// TIA Portal V19 export
FUNCTION_BLOCK "HEATING_PROCEES"   // FB14, LAD
TITLE = Heating
{ S7_Optimized_Access := 'TRUE' }
// stored: MemoryReserve 100, SetENOAutomatically false
   VAR_INPUT
      CHS_CFB : Bool;
      UCHS_CFB : Bool;
      CSV_CFB : Bool;
      HEAT_RUNNING : Bool;
      SELECT_CHWS : Bool;
      SELECT_CTS : Bool;
      SELECT_HWS : Bool;
      RUNNING : Bool;
      ESTOP : Bool;
      RESET : Bool;
      UCHWS : Bool;
      CHWS : Bool;
      CTS : Bool;
      HWS : Bool;
      HWS_OFB : Bool;
      CTS_OFB : Bool;
      CHWS_OFB : Bool;
      PUMP_RUN : Bool;
      SP : Real;
      PV : Real;
   END_VAR
   VAR_OUTPUT
      UCHWS_CMD : Bool;
      UCHWR_CMD : Bool;
      CHWS_CMD : Bool;
      CHWR_CMD : Bool;
      CTS_CMD : Bool;
      CTR_CMD : Bool;
      HWS_CMD : Bool;
      HWR_CMD : Bool;
      PUMP_CMD : Bool;
      CV_CMD : Bool;
   END_VAR
   VAR
      IEC_Timer_0_Instance : TP_TIME;
      IEC_Timer_1_Instance_1 { S7_SetPoint := 'True'} : TP_TIME;
      IEC_Timer_0_Instance_1 { S7_SetPoint := 'True'} : TP_TIME;
      IEC_Timer_0_Instance_2 { S7_SetPoint := 'True'} : TP_TIME;
      IEC_Timer_0_Instance_3 { S7_SetPoint := 'True'} : TP_TIME;
      IEC_Timer_0_Instance_4 { S7_SetPoint := 'True'} : TP_TIME;
      IEC_Timer_0_Instance_5 { S7_SetPoint := 'True'} : TP_TIME;
      IEC_Timer_0_Instance_6 { S7_SetPoint := 'True'} : TP_TIME;
      IEC_Timer_0_Instance_7 { S7_SetPoint := 'True'} : TP_TIME;
      IEC_Timer_0_Instance_8 { S7_SetPoint := 'True'} : TP_TIME;
      IEC_Timer_0_Instance_9 { S7_SetPoint := 'True'} : TP_TIME;
      "STEP" { S7_SetPoint := 'True'} : Int;
      P_TRIG : Bool;
      P_TRIG_1 : Bool;
      P_TRIG_2 : Bool;
      P_TRIG_3 : Bool;
      P_TRIG_4 : Bool;
      P_TRIG_5 : Bool;
      P_TRIG_6 : Bool;
      P_TRIG_7 : Bool;
      P_TRIG_8 : Bool;
      P_TRIG_9 : Bool;
      P_TRIG_10 : Bool;
      P_TRIG_11 : Bool;
      P_TRIG_12 : Bool;
      P_TRIG_13 : Bool;
      P_TRIG_14 : Bool;
      P_TRIG_15 : Bool;
      P_TRIG_16 : Bool;
      IEC_Timer_0_Instance_10 { S7_SetPoint := 'True'} : TP_TIME;
      IEC_Timer_0_Instance_11 { S7_SetPoint := 'True'} : TON_TIME;
      IEC_Timer_0_Instance_12 { S7_SetPoint := 'True'} : TON_TIME;
   END_VAR
   VAR_TEMP   // added for the SCL form of the ladder/FBD networks
      _w1 : Bool;
      _w2 : Bool;
      _w3 : Bool;
      _w4 : Bool;
      _w5 : Bool;
      _w6 : Bool;
      _w7 : Bool;
      _w8 : Bool;
   END_VAR
BEGIN

REGION Network 1: ULTRACHILLED TO CHILLED MODE
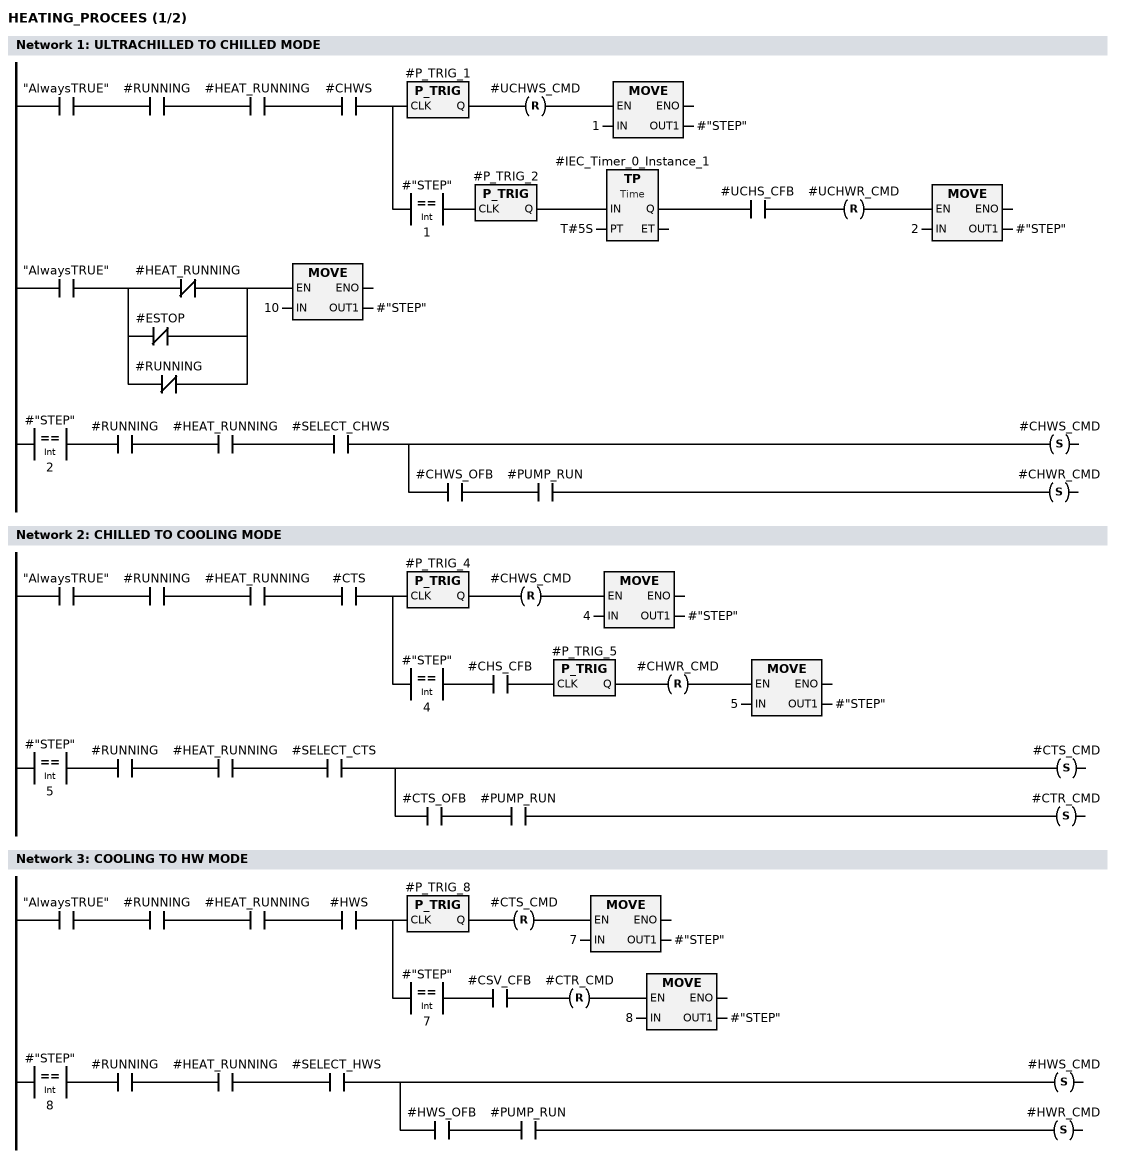
   RUNG wire#powerrail
      Contact( "AlwaysTRUE" )
      Contact( #RUNNING )
      Contact( #HEAT_RUNNING )
      Contact( #CHWS )
      wire#w1
      P_Trig( #P_TRIG_1 )
      R_Coil( #UCHWS_CMD )
      Move(in := 1, out1 => #"STEP")
   END_RUNG
   RUNG wire#w1
      { S7_Templates := "SrcType := Int" } EQ_Contact(in1 := #"STEP", in2 := 1)
      P_Trig( #P_TRIG_2 )
      { S7_Templates := "time_type := Time" } #IEC_Timer_0_Instance_1.TP(pt := T#5S, et =>)
      Contact( #UCHS_CFB )
      R_Coil( #UCHWR_CMD )
      Move(in := 2, out1 => #"STEP")
   END_RUNG
   RUNG wire#powerrail
      Contact( "AlwaysTRUE" )
      wire#w2
      I_Contact( #HEAT_RUNNING )
      wire#w3
      Move(in := 10, out1 => #"STEP")
   END_RUNG
   RUNG wire#w2
      I_Contact( #ESTOP )
   END_RUNG wire#w3
   RUNG wire#w2
      I_Contact( #RUNNING )
   END_RUNG wire#w3
   RUNG wire#powerrail
      { S7_Templates := "SrcType := Int" } EQ_Contact(in1 := #"STEP", in2 := 2)
      Contact( #RUNNING )
      Contact( #HEAT_RUNNING )
      Contact( #SELECT_CHWS )
      wire#w4
      S_Coil( #CHWS_CMD )
   END_RUNG
   RUNG wire#w4
      Contact( #CHWS_OFB )
      Contact( #PUMP_RUN )
      S_Coil( #CHWR_CMD )
   END_RUNG
   // the same network as SCL:
   #_w1 := "AlwaysTRUE" AND #RUNNING AND #HEAT_RUNNING AND #CHWS;
   #_w2 := #_w1 AND NOT #P_TRIG_1;   // rising edge
   #P_TRIG_1 := #_w1;
   IF #_w2 THEN
       #UCHWS_CMD := FALSE;
       #"STEP" := 1;
   END_IF;
   #_w3 := #_w1 AND (#"STEP" = 1);
   #_w4 := #_w3 AND NOT #P_TRIG_2;   // rising edge
   #P_TRIG_2 := #_w3;
   #IEC_Timer_0_Instance_1(IN := #_w4, PT := T#5S);   // TP
   IF #IEC_Timer_0_Instance_1.Q AND #UCHS_CFB THEN
       #UCHWR_CMD := FALSE;
       #"STEP" := 2;
   END_IF;
   IF "AlwaysTRUE" AND (NOT #HEAT_RUNNING OR NOT #ESTOP OR NOT #RUNNING) THEN #"STEP" := 10; END_IF;
   #_w5 := (#"STEP" = 2) AND #RUNNING AND #HEAT_RUNNING AND #SELECT_CHWS;
   IF #_w5 THEN #CHWS_CMD := TRUE; END_IF;
   IF #_w5 AND #CHWS_OFB AND #PUMP_RUN THEN #CHWR_CMD := TRUE; END_IF;
END_REGION

REGION Network 2: CHILLED TO COOLING MODE
   RUNG wire#powerrail
      Contact( "AlwaysTRUE" )
      Contact( #RUNNING )
      Contact( #HEAT_RUNNING )
      Contact( #CTS )
      wire#w1
      P_Trig( #P_TRIG_4 )
      R_Coil( #CHWS_CMD )
      Move(in := 4, out1 => #"STEP")
   END_RUNG
   RUNG wire#w1
      { S7_Templates := "SrcType := Int" } EQ_Contact(in1 := #"STEP", in2 := 4)
      Contact( #CHS_CFB )
      P_Trig( #P_TRIG_5 )
      R_Coil( #CHWR_CMD )
      Move(in := 5, out1 => #"STEP")
   END_RUNG
   RUNG wire#powerrail
      { S7_Templates := "SrcType := Int" } EQ_Contact(in1 := #"STEP", in2 := 5)
      Contact( #RUNNING )
      Contact( #HEAT_RUNNING )
      Contact( #SELECT_CTS )
      wire#w2
      S_Coil( #CTS_CMD )
   END_RUNG
   RUNG wire#w2
      Contact( #CTS_OFB )
      Contact( #PUMP_RUN )
      S_Coil( #CTR_CMD )
   END_RUNG
   // the same network as SCL:
   #_w1 := "AlwaysTRUE" AND #RUNNING AND #HEAT_RUNNING AND #CTS;
   #_w2 := #_w1 AND NOT #P_TRIG_4;   // rising edge
   #P_TRIG_4 := #_w1;
   IF #_w2 THEN
       #CHWS_CMD := FALSE;
       #"STEP" := 4;
   END_IF;
   #_w3 := #_w1 AND (#"STEP" = 4) AND #CHS_CFB;
   #_w4 := #_w3 AND NOT #P_TRIG_5;   // rising edge
   #P_TRIG_5 := #_w3;
   IF #_w4 THEN
       #CHWR_CMD := FALSE;
       #"STEP" := 5;
   END_IF;
   #_w5 := (#"STEP" = 5) AND #RUNNING AND #HEAT_RUNNING AND #SELECT_CTS;
   IF #_w5 THEN #CTS_CMD := TRUE; END_IF;
   IF #_w5 AND #CTS_OFB AND #PUMP_RUN THEN #CTR_CMD := TRUE; END_IF;
END_REGION

REGION Network 3: COOLING TO HW MODE
   RUNG wire#powerrail
      Contact( "AlwaysTRUE" )
      Contact( #RUNNING )
      Contact( #HEAT_RUNNING )
      Contact( #HWS )
      wire#w1
      P_Trig( #P_TRIG_8 )
      R_Coil( #CTS_CMD )
      Move(in := 7, out1 => #"STEP")
   END_RUNG
   RUNG wire#w1
      { S7_Templates := "SrcType := Int" } EQ_Contact(in1 := #"STEP", in2 := 7)
      Contact( #CSV_CFB )
      R_Coil( #CTR_CMD )
      Move(in := 8, out1 => #"STEP")
   END_RUNG
   RUNG wire#powerrail
      { S7_Templates := "SrcType := Int" } EQ_Contact(in1 := #"STEP", in2 := 8)
      Contact( #RUNNING )
      Contact( #HEAT_RUNNING )
      Contact( #SELECT_HWS )
      wire#w2
      S_Coil( #HWS_CMD )
   END_RUNG
   RUNG wire#w2
      Contact( #HWS_OFB )
      Contact( #PUMP_RUN )
      S_Coil( #HWR_CMD )
   END_RUNG
   // the same network as SCL:
   #_w1 := "AlwaysTRUE" AND #RUNNING AND #HEAT_RUNNING AND #HWS;
   #_w2 := #_w1 AND NOT #P_TRIG_8;   // rising edge
   #P_TRIG_8 := #_w1;
   IF #_w2 THEN
       #CTS_CMD := FALSE;
       #"STEP" := 7;
   END_IF;
   IF #_w1 AND (#"STEP" = 7) AND #CSV_CFB THEN
       #CTR_CMD := FALSE;
       #"STEP" := 8;
   END_IF;
   #_w3 := (#"STEP" = 8) AND #RUNNING AND #HEAT_RUNNING AND #SELECT_HWS;
   IF #_w3 THEN #HWS_CMD := TRUE; END_IF;
   IF #_w3 AND #HWS_OFB AND #PUMP_RUN THEN #HWR_CMD := TRUE; END_IF;
END_REGION

REGION Network 4
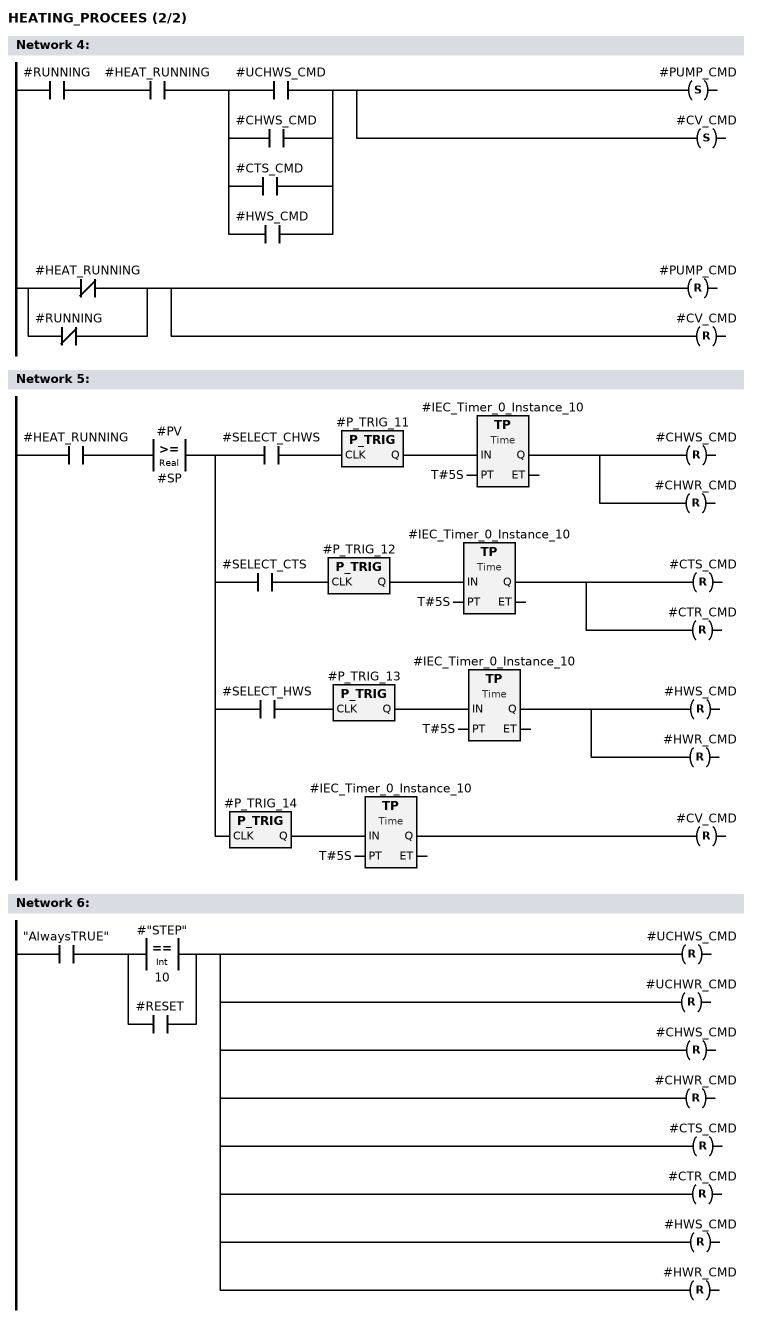
   RUNG wire#powerrail
      Contact( #RUNNING )
      Contact( #HEAT_RUNNING )
      wire#w1
      Contact( #UCHWS_CMD )
      wire#w2
      S_Coil( #PUMP_CMD )
   END_RUNG
   RUNG wire#w1
      Contact( #CHWS_CMD )
   END_RUNG wire#w2
   RUNG wire#w1
      Contact( #CTS_CMD )
   END_RUNG wire#w2
   RUNG wire#w1
      Contact( #HWS_CMD )
   END_RUNG wire#w2
   RUNG wire#w2
      S_Coil( #CV_CMD )
   END_RUNG
   RUNG wire#powerrail
      I_Contact( #HEAT_RUNNING )
      wire#w3
      R_Coil( #PUMP_CMD )
   END_RUNG
   RUNG wire#powerrail
      I_Contact( #RUNNING )
   END_RUNG wire#w3
   RUNG wire#w3
      R_Coil( #CV_CMD )
   END_RUNG
   // the same network as SCL:
   IF #RUNNING AND #HEAT_RUNNING AND (#UCHWS_CMD OR #CHWS_CMD OR #CTS_CMD OR #HWS_CMD) THEN
       #PUMP_CMD := TRUE;
       #CV_CMD := TRUE;
   END_IF;
   IF NOT #HEAT_RUNNING OR NOT #RUNNING THEN
       #PUMP_CMD := FALSE;
       #CV_CMD := FALSE;
   END_IF;
END_REGION

REGION Network 5
   RUNG wire#powerrail
      Contact( #HEAT_RUNNING )
      { S7_Templates := "SrcType := Real" } GE_Contact(in1 := #PV, in2 := #SP)
      wire#w1
      Contact( #SELECT_CHWS )
      P_Trig( #P_TRIG_11 )
      { S7_Templates := "time_type := Time" } #IEC_Timer_0_Instance_10.TP(pt := T#5S, et =>)
      wire#w2
      R_Coil( #CHWS_CMD )
   END_RUNG
   RUNG wire#w2
      R_Coil( #CHWR_CMD )
   END_RUNG
   RUNG wire#w1
      Contact( #SELECT_CTS )
      P_Trig( #P_TRIG_12 )
      { S7_Templates := "time_type := Time" } #IEC_Timer_0_Instance_10.TP(pt := T#5S, et =>)
      wire#w3
      R_Coil( #CTS_CMD )
   END_RUNG
   RUNG wire#w3
      R_Coil( #CTR_CMD )
   END_RUNG
   RUNG wire#w1
      Contact( #SELECT_HWS )
      P_Trig( #P_TRIG_13 )
      { S7_Templates := "time_type := Time" } #IEC_Timer_0_Instance_10.TP(pt := T#5S, et =>)
      wire#w4
      R_Coil( #HWS_CMD )
   END_RUNG
   RUNG wire#w4
      R_Coil( #HWR_CMD )
   END_RUNG
   RUNG wire#w1
      P_Trig( #P_TRIG_14 )
      { S7_Templates := "time_type := Time" } #IEC_Timer_0_Instance_10.TP(pt := T#5S, et =>)
      R_Coil( #CV_CMD )
   END_RUNG
   // the same network as SCL:
   #_w1 := #HEAT_RUNNING AND (#PV >= #SP);
   #_w2 := #_w1 AND #SELECT_CHWS;
   #_w3 := #_w2 AND NOT #P_TRIG_11;   // rising edge
   #P_TRIG_11 := #_w2;
   #IEC_Timer_0_Instance_10(IN := #_w3, PT := T#5S);   // TP
   IF #IEC_Timer_0_Instance_10.Q THEN
       #CHWS_CMD := FALSE;
       #CHWR_CMD := FALSE;
   END_IF;
   #_w4 := #_w1 AND #SELECT_CTS;
   #_w5 := #_w4 AND NOT #P_TRIG_12;   // rising edge
   #P_TRIG_12 := #_w4;
   #IEC_Timer_0_Instance_10(IN := #_w5, PT := T#5S);   // TP
   IF #IEC_Timer_0_Instance_10.Q THEN
       #CTS_CMD := FALSE;
       #CTR_CMD := FALSE;
   END_IF;
   #_w6 := #_w1 AND #SELECT_HWS;
   #_w7 := #_w6 AND NOT #P_TRIG_13;   // rising edge
   #P_TRIG_13 := #_w6;
   #IEC_Timer_0_Instance_10(IN := #_w7, PT := T#5S);   // TP
   IF #IEC_Timer_0_Instance_10.Q THEN
       #HWS_CMD := FALSE;
       #HWR_CMD := FALSE;
   END_IF;
   #_w8 := #_w1 AND NOT #P_TRIG_14;   // rising edge
   #P_TRIG_14 := #_w1;
   #IEC_Timer_0_Instance_10(IN := #_w8, PT := T#5S);   // TP
   IF #IEC_Timer_0_Instance_10.Q THEN #CV_CMD := FALSE; END_IF;
END_REGION

REGION Network 6
   RUNG wire#powerrail
      Contact( "AlwaysTRUE" )
      wire#w1
      { S7_Templates := "SrcType := Int" } EQ_Contact(in1 := #"STEP", in2 := 10)
      wire#w2
      R_Coil( #UCHWS_CMD )
   END_RUNG
   RUNG wire#w1
      Contact( #RESET )
   END_RUNG wire#w2
   RUNG wire#w2
      R_Coil( #UCHWR_CMD )
   END_RUNG
   RUNG wire#w2
      R_Coil( #CHWS_CMD )
   END_RUNG
   RUNG wire#w2
      R_Coil( #CHWR_CMD )
   END_RUNG
   RUNG wire#w2
      R_Coil( #CTS_CMD )
   END_RUNG
   RUNG wire#w2
      R_Coil( #CTR_CMD )
   END_RUNG
   RUNG wire#w2
      R_Coil( #HWS_CMD )
   END_RUNG
   RUNG wire#w2
      R_Coil( #HWR_CMD )
   END_RUNG
   // the same network as SCL:
   IF "AlwaysTRUE" AND ((#"STEP" = 10) OR #RESET) THEN
       #UCHWS_CMD := FALSE;
       #UCHWR_CMD := FALSE;
       #CHWS_CMD := FALSE;
       #CHWR_CMD := FALSE;
       #CTS_CMD := FALSE;
       #CTR_CMD := FALSE;
       #HWS_CMD := FALSE;
       #HWR_CMD := FALSE;
   END_IF;
END_REGION
END_FUNCTION_BLOCK
